Fanuc KAREL source: kt00751.KL

-- PROVISIONAL review KL for V1013-1; original PC SHA256 5007599ea7ab6464150a4f547bb08dfd2407cb59cbe77610e4ad61ea5f5c867a
-- Incomplete behavior may be omitted. Consult companion uncertainty JSON. Do not deploy.
PROGRAM KT00751
%NOLOCKGROUP
VAR
  R1 : REAL
  R2 : REAL
  OUT : REAL
BEGIN
  -- UNRESOLVED_PC offsets 5-16; opcodes 2E,23
  -- UNRESOLVED_PC offsets 21-32; opcodes 2E,23
  -- UNRESOLVED_PC offsets 37-48; opcodes 2E,23
  -- UNRESOLVED_PC offsets 53-64; opcodes 2E,23
  -- UNRESOLVED_PC offsets 69-82; opcodes 21,67,23
  -- UNRESOLVED_PC offsets 87-91; opcodes 7F
END KT00751
